(* IEC 61131-3 sources: nautilus/examples/remote-fleet/sites/well-1, 3 files *)

(* ---- types.st ---- *)
(* A root .st file with no PROGRAM is a project library, in scope for
   every task's compile — see docs/functions.md "A .ld library" (the same
   rule, one language over). Pump is the SAME shape scada/sites.yaml
   declares as its shared Template for all three sites, but this copy, not
   a shared package, is what ships: each site deploys alone. *)
TYPE
  Pump : STRUCT
    Run     : BOOL;   (* running feedback *)
    Fault   : BOOL;   (* VFD fault *)
    SpeedHz : LREAL;  (* actual speed *)
    SpeedSP : LREAL;  (* operator/SCADA setpoint — written locally or by
                         a Sparkplug NCMD member write from the SCADA host *)
  END_STRUCT;
END_TYPE

(* ---- sim.st ---- *)
(* Bench-only plant: the wet well's level (an inflow/outflow balance) and
   the pump/VFD's speed response. A field deployment deletes this task
   and points well.st's Pump1/WellLevel tags at real hardware instead
   (a Modbus VFD and level transmitter — see ../booster-1/devices.yaml
   for the pattern this fleet uses elsewhere). *)
PROGRAM Sim
VAR_EXTERNAL
    WellLevel      : LREAL;
    InflowLps      : LREAL;
    Pump1          : Pump;
    Pump1_RunCmd   : BOOL;
    Pump1_SpeedCmd : LREAL;
    SimDtS         : LREAL;
END_VAR
VAR
    outflowLps : LREAL;
    tSec       : LREAL;
END_VAR
VAR CONSTANT
    InflowVaryFrac : LREAL := 0.20;
    InflowPeriodS  : LREAL := 180.0;
    TwoPi          : LREAL := 6.2831853;
END_VAR

tSec := tSec + SimDtS;

(* Speed ramps toward the command at 10 Hz/s; running is "spinning". *)
IF Pump1_RunCmd THEN
    Pump1.SpeedHz := LIMIT(0.0, Pump1.SpeedHz + LIMIT(-10.0 * SimDtS, Pump1_SpeedCmd - Pump1.SpeedHz, 10.0 * SimDtS), 60.0);
ELSE
    Pump1.SpeedHz := MAX(0.0, Pump1.SpeedHz - 10.0 * SimDtS);
END_IF;
Pump1.Run := Pump1.SpeedHz > 5.0;
Pump1.Fault := FALSE;

(* Discharge flow: ~0 below 25 Hz, 10 L/s at 60 Hz, linear between — a
   small well pump, a tenth the size of lift-station's lift pumps. *)
IF Pump1.SpeedHz <= 25.0 THEN
    outflowLps := 0.0;
ELSE
    outflowLps := (Pump1.SpeedHz - 25.0) / (60.0 - 25.0) * 10.0;
END_IF;

(* 1500 L span over 100 % (15 L per %) plus a slow sinusoid on the base
   inflow, so the level never sits dead flat. *)
WellLevel := LIMIT(0.0, WellLevel + (InflowLps * (1.0 + InflowVaryFrac * SIN(tSec / InflowPeriodS * TwoPi)) - outflowLps) * SimDtS / 15.0, 100.0);
END_PROGRAM

(* ---- well.st ---- *)
(* well-1's own control: a single pump, called on rising wet-well level
   with hysteresis, run at a speed clamped to [MinSpeedHz, MaxSpeedHz].
   Pump1 is a Sparkplug Template (TYPE Pump, types.st) — the SAME shape
   scada/sites.yaml declares for all three sites, but this file, not a
   shared library, is where it lives: each site deploys alone (see
   ../../README.md). *)
PROGRAM Well
VAR_EXTERNAL
    WellLevel     : LREAL;
    Pump1         : Pump;
    Pump1_RunCmd  : BOOL;
    Pump1_SpeedCmd : LREAL;
    PumpOnLevel   : LREAL;
    PumpOffLevel  : LREAL;
    MinSpeedHz    : LREAL;
    MaxSpeedHz    : LREAL;
    PumpStarts    : INT;
    PumpHours     : LREAL;
    WellDtS       : LREAL;
END_VAR
VAR
    edgeUp : R_TRIG;
END_VAR

(* Seal-in hysteresis: call the pump at PumpOnLevel, hold it until the
   level drops back through PumpOffLevel — same idiom as lift-station's
   HighLevelAlm seal-in, one line instead of a state machine. *)
Pump1_RunCmd := (WellLevel >= PumpOnLevel) OR (Pump1_RunCmd AND WellLevel > PumpOffLevel);

IF Pump1_RunCmd THEN
    Pump1_SpeedCmd := LIMIT(MinSpeedHz, Pump1.SpeedSP, MaxSpeedHz);
ELSE
    Pump1_SpeedCmd := 0.0;
END_IF;

(* Run-hours meter: starts on Run's rising edge, hours while running. *)
edgeUp(CLK := Pump1.Run);
IF edgeUp.Q THEN
    PumpStarts := PumpStarts + 1;
END_IF;
IF Pump1.Run THEN
    PumpHours := PumpHours + WellDtS / 3600.0;
END_IF;
END_PROGRAM
